Fanuc KAREL source: KT00781.KL

PROGRAM KT00781
%NOLOCKGROUP
VAR
  B1: BOOLEAN
  B2: BOOLEAN
  OUT: REAL
BEGIN
  B1 = TRUE
  B2 = FALSE
  B1 = TRUE
  B2 = FALSE
  OUT = ASIN(B1)
END KT00781
